Staubli VAL3: safeData.pjx

--- safeData.pjx ---
Parameters version=s8.10.3Cs9_BS2093 stackSize=5000 millimeterUnit=true
Program file=start.pgx
Program file=stop.pgx
Data file=safeData.dtx
Type name=zoneItem path=Disk://source/template/zoneTemplate/zoneTemplate.pjx
Type name=sPoint path=Disk://source/template/sPointTemplate/sPointTemplate.pjx

--- safeData.dtx ---
public sPoint sSPoint[10]
  [0]
    bool bActive
    pointRx pPointRx = {x=108.485671, y=75.476203, z=519.0997746, rx=-0.682186, ry=-2.964024, rz=96.292694, shoulder=lefty, elbow=enegative, wrist=wpositive, fatherId=world[0]}
    string sName = "安全点0"
  [1]
    bool bActive = true
    pointRx pPointRx = {x=1213.921571, y=199.805628, z=237.299989, rx=14.382647, ry=120.0425711, rz=-19.201374, shoulder=lefty, elbow=epositive, wrist=wpositive, fatherId=world[0]}
    string sName = "安全点1"
  [2]
    bool bActive
    pointRx pPointRx
    string sName = "安全点2"
  [3]
    bool bActive
    pointRx pPointRx
    string sName = "安全点3"
  [4]
    bool bActive
    pointRx pPointRx
    string sName = "安全点4"
  [5]
    bool bActive
    pointRx pPointRx
    string sName = "安全点5"
  [6]
    bool bActive
    pointRx pPointRx
    string sName = "安全点6"
  [7]
    bool bActive
    pointRx pPointRx
    string sName = "安全点7"
  [8]
    bool bActive
    pointRx pPointRx
    string sName = "安全点8"
  [9]
    bool bActive
    pointRx pPointRx
    string sName = "安全点9"
public zoneItem zZoneItem[10]
  [0]
    bool bActive = true
    frame fBase
    pointRx pFirst = {x=108.485671, y=75.476203, z=519.0997746, rx=-0.682186, ry=-2.964024, rz=96.292694, shoulder=lefty, elbow=enegative, wrist=wpositive}
    pointRx pO
    pointRx pSecond = {x=500, y=500, z=500}
    pointRx pX
    pointRx pY
    string sID = "rrff"
  [1]
    bool bActive
    frame fBase
    pointRx pFirst
    pointRx pO
    pointRx pSecond
    pointRx pX
    pointRx pY
    string sID = "干涉区1"
  [2]
    bool bActive
    frame fBase
    pointRx pFirst
    pointRx pO
    pointRx pSecond
    pointRx pX
    pointRx pY
    string sID = "干涉区2"
  [3]
    bool bActive
    frame fBase
    pointRx pFirst
    pointRx pO
    pointRx pSecond
    pointRx pX
    pointRx pY
    string sID = "干涉区3"
  [4]
    bool bActive
    frame fBase
    pointRx pFirst
    pointRx pO
    pointRx pSecond
    pointRx pX
    pointRx pY
    string sID = "干涉区4"
  [5]
    bool bActive
    frame fBase
    pointRx pFirst
    pointRx pO
    pointRx pSecond
    pointRx pX
    pointRx pY
    string sID = "干涉区5"
  [6]
    bool bActive
    frame fBase
    pointRx pFirst
    pointRx pO
    pointRx pSecond
    pointRx pX
    pointRx pY
    string sID = "干涉区6"
  [7]
    bool bActive
    frame fBase
    pointRx pFirst
    pointRx pO
    pointRx pSecond
    pointRx pX
    pointRx pY
    string sID = "干涉区7"
  [8]
    bool bActive
    frame fBase
    pointRx pFirst
    pointRx pO
    pointRx pSecond
    pointRx pX
    pointRx pY
    string sID = "干涉区8"
  [9]
    bool bActive
    frame fBase
    pointRx pFirst
    pointRx pO
    pointRx pSecond
    pointRx pX
    pointRx pY
    string sID = "干涉区9"

--- start.pgx ---
program start()
begin
end

--- stop.pgx ---
program stop()
begin
end
